(* IEC 61131-3 sources: bevling_machine/framework/sources/03_Units, 8 files *)

(* ---- FB_ClearanceUnit.st ---- *)
(* 模块说明：并行执行 P/Q 两路避让；两路都完成才继续，任一路故障向主流程报告。 *)
FUNCTION_BLOCK FB_ClearanceUnit
VAR_INPUT
    xExecute : BOOL; (* 子流程执行许可；须保持到完成，清 FALSE 复位该流程步骤和错误。 *)
    stRecipe : ST_Recipe; (* 待校验配方或上层传入的运行配方，字段含义见 ST_Recipe。 *)
END_VAR
VAR_IN_OUT
    aCommand : ARRAY[1..17] OF ST_DeviceCommand; (* 统一设备请求数组 1..17；子流程写请求，设备管理器执行。 *)
    aStatus : ARRAY[1..17] OF ST_DeviceStatus; (* 各设备的反馈数组 1..17，供判断忙、完成序号、故障和位置。 *)
    udiCounter : UDINT; (* 全机共享的动作序号计数器，通过引用传递；由 F_NextID 分配，0 不使用。 *)
END_VAR
VAR_OUTPUT
    xDone : BOOL; (* 本子流程完成标志；执行许可撤销后复位。 *)
    xError : BOOL; (* 本设备或本子流程发生故障；具体原因见对应错误码。 *)
    udiErrorID : UDINT; (* 错误码；0 表示无错误，设备或流程发生异常时赋值。 *)
    uiLengthStep : UINT; (* 定长支线当前步骤，供监控定位等待点。 *)
    uiTransferStep : UINT; (* 流利条/侧推/侧挡支线当前步骤，供监控定位等待点。 *)
END_VAR
VAR
    fbLength : FB_ClearLength; (* P 支线：D5 升起、D4 移开。 *)
    fbTransfer : FB_ClearTransfer; (* 切割前流利条/侧推/侧挡避让支线。 *)
END_VAR
FUNCTION_BLOCK FB_ClearanceUnit
(* P/Q 两路同一扫描使能；xDone 使用 AND，任一路未完成均不得继续。 *)
fbLength(xExecute:=xExecute,stRecipe:=stRecipe,aCommand:=aCommand,aStatus:=aStatus,udiCounter:=udiCounter);
fbTransfer(xExecute:=xExecute,stRecipe:=stRecipe,aCommand:=aCommand,aStatus:=aStatus,udiCounter:=udiCounter);
xDone := fbLength.xDone AND fbTransfer.xDone;
xError := fbLength.xError OR fbTransfer.xError;
udiErrorID := MAX(fbLength.udiErrorID,fbTransfer.udiErrorID);
uiLengthStep := fbLength.uiStep; uiTransferStep := fbTransfer.uiStep;

(* ---- FB_ClearLength.st ---- *)
(* 模块说明：切割前避让支线 P：D5 定长升起，再将 D4 移到避让位置。每步等待本次序号完成。 *)
FUNCTION_BLOCK FB_ClearLength
VAR_INPUT
    xExecute : BOOL; (* 子流程执行许可；须保持到完成，清 FALSE 复位该流程步骤和错误。 *)
    stRecipe : ST_Recipe; (* 待校验配方或上层传入的运行配方，字段含义见 ST_Recipe。 *)
END_VAR
VAR_IN_OUT
    aCommand : ARRAY[1..17] OF ST_DeviceCommand; (* 统一设备请求数组 1..17；子流程写请求，设备管理器执行。 *)
    aStatus : ARRAY[1..17] OF ST_DeviceStatus; (* 各设备的反馈数组 1..17，供判断忙、完成序号、故障和位置。 *)
    udiCounter : UDINT; (* 全机共享的动作序号计数器，通过引用传递；由 F_NextID 分配，0 不使用。 *)
END_VAR
VAR_OUTPUT
    xDone : BOOL; (* 本子流程完成标志；执行许可撤销后复位。 *)
    xError : BOOL; (* 本设备或本子流程发生故障；具体原因见对应错误码。 *)
    udiErrorID : UDINT; (* 非法步骤码 4100；动作超时码=4100+uiStep，可据此定位本支线等待点。 *)
    uiStep : UINT; (* 当前子步骤：0 待机，10/20/... 执行动作，1000 完成；切勿在线强制跳步。 *)
END_VAR
VAR
    uiPrevStep : UINT := 65535; (* 上扫描步骤，用于判断本扫描是否刚进入新步骤。 *)
    udiToken : UDINT; (* 本步骤专用动作序号；同一步中的设备共用该号，以排除旧完成信号。 *)
    xEntry : BOOL; (* 本扫描为新步骤入口；用于分配新序号并复位步骤超时计时。 *)
    tonStep : TON; (* 步骤超时定时器；进入新步骤时复位，超时错误码由模块及当前步号组成。 *)
    tonSpray : TON; (* 通用子流程模板的喷油定时器，只有 FB_ReturnKnife 用其完成条件。 *)
END_VAR
FUNCTION_BLOCK FB_ClearLength
(* 执行许可撤销即复位；步骤入口换新序号，每步等待本次动作完成，超时码=模块基码+步号。 *)
IF NOT xExecute THEN uiStep := 0; xError := FALSE; udiErrorID := 0; END_IF;
xEntry := uiStep <> uiPrevStep;
IF xEntry THEN udiToken := F_NextID(udiCounter); END_IF;
uiPrevStep := uiStep;
tonStep(IN := xExecute AND (uiStep > 0) AND (uiStep < 1000) AND NOT xEntry, PT := stRecipe.tStepTimeout);
tonSpray(IN := xExecute AND (uiStep = 10) AND aStatus[13].xActive, PT := stRecipe.tSpray);
IF xExecute AND NOT xError THEN
CASE uiStep OF
0: (* 待机；许可有效时进入首个动作。 *) uiStep := 10;
10: (* P010 定长 D5 升起避让；确认本次动作完成后再允许 D4 平移。 *)
aCommand[5] := F_Command(E_DeviceAction.Position, udiToken, 0.0, stRecipe.lrPositionVelocity);
IF F_Done(aStatus[5], udiToken) THEN uiStep := 20; END_IF;
20: (* P020 定长 D4 移到配方避让位置，等待本次序号完成。 *)
aCommand[4] := F_Command(E_DeviceAction.Position, udiToken, stRecipe.lrLengthClear, stRecipe.lrPositionVelocity);
IF F_Done(aStatus[4], udiToken) THEN uiStep := 1000; END_IF;
1000: (* 本支线完成，保持至 xExecute 撤销。 *) ;
ELSE xError := TRUE; udiErrorID := 4100;
END_CASE;
IF tonStep.Q THEN xError := TRUE; udiErrorID := 4100 + UINT_TO_UDINT(uiStep); END_IF;
END_IF;
xDone := xExecute AND (uiStep = 1000) AND NOT xError;

(* ---- FB_ClearTransfer.st ---- *)
(* 模块说明：切割前避让支线 Q：G4 流利条下降、G3 解除侧推、G2 侧挡下降。 *)
FUNCTION_BLOCK FB_ClearTransfer
VAR_INPUT
    xExecute : BOOL; (* 子流程执行许可；须保持到完成，清 FALSE 复位该流程步骤和错误。 *)
    stRecipe : ST_Recipe; (* 待校验配方或上层传入的运行配方，字段含义见 ST_Recipe。 *)
END_VAR
VAR_IN_OUT
    aCommand : ARRAY[1..17] OF ST_DeviceCommand; (* 统一设备请求数组 1..17；子流程写请求，设备管理器执行。 *)
    aStatus : ARRAY[1..17] OF ST_DeviceStatus; (* 各设备的反馈数组 1..17，供判断忙、完成序号、故障和位置。 *)
    udiCounter : UDINT; (* 全机共享的动作序号计数器，通过引用传递；由 F_NextID 分配，0 不使用。 *)
END_VAR
VAR_OUTPUT
    xDone : BOOL; (* 本子流程完成标志；执行许可撤销后复位。 *)
    xError : BOOL; (* 本设备或本子流程发生故障；具体原因见对应错误码。 *)
    udiErrorID : UDINT; (* 非法步骤码 4200；动作超时码=4200+uiStep，可据此定位本支线等待点。 *)
    uiStep : UINT; (* 当前子步骤：0 待机，10/20/... 执行动作，1000 完成；切勿在线强制跳步。 *)
END_VAR
VAR
    uiPrevStep : UINT := 65535; (* 上扫描步骤，用于判断本扫描是否刚进入新步骤。 *)
    udiToken : UDINT; (* 本步骤专用动作序号；同一步中的设备共用该号，以排除旧完成信号。 *)
    xEntry : BOOL; (* 本扫描为新步骤入口；用于分配新序号并复位步骤超时计时。 *)
    tonStep : TON; (* 步骤超时定时器；进入新步骤时复位，超时错误码由模块及当前步号组成。 *)
    tonSpray : TON; (* 通用子流程模板的喷油定时器，只有 FB_ReturnKnife 用其完成条件。 *)
END_VAR
FUNCTION_BLOCK FB_ClearTransfer
(* 执行许可撤销即复位；步骤入口换新序号，每步等待本次动作完成，超时码=模块基码+步号。 *)
IF NOT xExecute THEN uiStep := 0; xError := FALSE; udiErrorID := 0; END_IF;
xEntry := uiStep <> uiPrevStep;
IF xEntry THEN udiToken := F_NextID(udiCounter); END_IF;
uiPrevStep := uiStep;
tonStep(IN := xExecute AND (uiStep > 0) AND (uiStep < 1000) AND NOT xEntry, PT := stRecipe.tStepTimeout);
tonSpray(IN := xExecute AND (uiStep = 10) AND aStatus[13].xActive, PT := stRecipe.tSpray);
IF xExecute AND NOT xError THEN
CASE uiStep OF
0: (* 待机；许可有效时进入首个动作。 *) uiStep := 10;
10: (* Q010 流利条 G4 下降。 *)
aCommand[12] := F_Command(E_DeviceAction.Position, udiToken, 0.0, stRecipe.lrPositionVelocity);
IF F_Done(aStatus[12], udiToken) THEN uiStep := 20; END_IF;
20: (* Q020 推动气缸 G3 放开。 *)
aCommand[11] := F_Command(E_DeviceAction.Position, udiToken, 0.0, stRecipe.lrPositionVelocity);
IF F_Done(aStatus[11], udiToken) THEN uiStep := 30; END_IF;
30: (* Q030 侧挡 G2 下降。目标固定发 1.0：本层不知道侧挡是单缸还是 300/450/600 三缸组，
   由设备层自己解释——仿真气缸按 1.0 到伸出端，真实三缸组按当前料型选缸下降。 *)
aCommand[10] := F_Command(E_DeviceAction.Position, udiToken, 1.0, stRecipe.lrPositionVelocity);
IF F_Done(aStatus[10], udiToken) THEN uiStep := 1000; END_IF;
1000: (* 本支线完成，保持至 xExecute 撤销。 *) ;
ELSE xError := TRUE; udiErrorID := 4200;
END_CASE;
IF tonStep.Q THEN xError := TRUE; udiErrorID := 4200 + UINT_TO_UDINT(uiStep); END_IF;
END_IF;
xDone := xExecute AND (uiStep = 1000) AND NOT xError;

(* ---- FB_Initialize.st ---- *)
(* 模块说明：初始姿态整理流程。20 步摆好避让姿态后，25 步让真实轴回零，30 步再按配方绝对定位。 *)
FUNCTION_BLOCK FB_Initialize
VAR_INPUT
    xExecute : BOOL; (* 子流程执行许可；须保持到完成，清 FALSE 复位该流程步骤和错误。 *)
    stRecipe : ST_Recipe; (* 待校验配方或上层传入的运行配方，字段含义见 ST_Recipe。 *)
END_VAR
VAR_IN_OUT
    aCommand : ARRAY[1..17] OF ST_DeviceCommand; (* 统一设备请求数组 1..17；子流程写请求，设备管理器执行。 *)
    aStatus : ARRAY[1..17] OF ST_DeviceStatus; (* 各设备的反馈数组 1..17，供判断忙、完成序号、故障和位置。 *)
    udiCounter : UDINT; (* 全机共享的动作序号计数器，通过引用传递；由 F_NextID 分配，0 不使用。 *)
END_VAR
VAR_OUTPUT
    xDone : BOOL; (* 本子流程完成标志；执行许可撤销后复位。 *)
    xError : BOOL; (* 本设备或本子流程发生故障；具体原因见对应错误码。 *)
    udiErrorID : UDINT; (* 非法步骤码 4600；动作超时码=4600+uiStep，可据此定位本支线等待点。 *)
    uiStep : UINT; (* 当前子步骤：0 待机，10/20/25/30/40 执行动作，1000 完成；切勿在线强制跳步。 *)
END_VAR
VAR
    uiPrevStep : UINT := 65535; (* 上扫描步骤，用于判断本扫描是否刚进入新步骤。 *)
    udiToken : UDINT; (* 本步骤专用动作序号；同一步中的设备共用该号，以排除旧完成信号。 *)
    xEntry : BOOL; (* 本扫描为新步骤入口；用于分配新序号并复位步骤超时计时。 *)
    tonStep : TON; (* 步骤超时定时器；进入新步骤时复位，超时错误码由模块及当前步号组成。 *)
    tonSpray : TON; (* 通用子流程模板的喷油定时器，只有 FB_ReturnKnife 用其完成条件。 *)
END_VAR
FUNCTION_BLOCK FB_Initialize
(* 执行许可撤销即复位；步骤入口换新序号，每步等待本次动作完成，超时码=模块基码+步号。 *)
IF NOT xExecute THEN uiStep := 0; xError := FALSE; udiErrorID := 0; END_IF;
xEntry := uiStep <> uiPrevStep;
IF xEntry THEN udiToken := F_NextID(udiCounter); END_IF;
uiPrevStep := uiStep;
tonStep(IN := xExecute AND (uiStep > 0) AND (uiStep < 1000) AND NOT xEntry, PT := stRecipe.tStepTimeout);
tonSpray(IN := xExecute AND (uiStep = 10) AND aStatus[13].xActive, PT := stRecipe.tSpray);
IF xExecute AND NOT xError THEN
CASE uiStep OF
0: (* 待机；许可有效时进入首个动作。 *) uiStep := 10;
10: (* 仿真初始化 10：同时抬起 G9、抬起 G1、打开 G8，三项都完成才继续。 *)
aCommand[17] := F_Command(E_DeviceAction.Position, udiToken, 0.0, stRecipe.lrPositionVelocity);
aCommand[9] := F_Command(E_DeviceAction.Position, udiToken, 0.0, stRecipe.lrPositionVelocity);
aCommand[16] := F_Command(E_DeviceAction.Position, udiToken, 0.0, stRecipe.lrPositionVelocity);
IF F_Done(aStatus[17], udiToken) AND F_Done(aStatus[9], udiToken) AND F_Done(aStatus[16], udiToken) THEN uiStep := 20; END_IF;
20: (* 仿真初始化 20：D5 升起、G2 提升、G3 释放、G4 提升、G7 下降，全部完成再定位。 *)
aCommand[5] := F_Command(E_DeviceAction.Position, udiToken, 0.0, stRecipe.lrPositionVelocity);
aCommand[10] := F_Command(E_DeviceAction.Position, udiToken, 0.0, stRecipe.lrPositionVelocity);
aCommand[11] := F_Command(E_DeviceAction.Position, udiToken, 0.0, stRecipe.lrPositionVelocity);
aCommand[12] := F_Command(E_DeviceAction.Position, udiToken, 1.0, stRecipe.lrPositionVelocity);
aCommand[15] := F_Command(E_DeviceAction.Position, udiToken, 0.0, stRecipe.lrPositionVelocity);
IF F_Done(aStatus[5], udiToken) AND F_Done(aStatus[10], udiToken) AND F_Done(aStatus[11], udiToken) AND F_Done(aStatus[12], udiToken) AND F_Done(aStatus[15], udiToken) THEN uiStep := 25; END_IF;
25: (* 初始化 25：真实轴回零。D2 走刀与 D8 旋转是真轴，D4 定长平移当前为仿真，由仿真在 tSimAction 后完成。
       D3 盘刀是连续旋转主轴，自动流程只下发 Run 不定位，因此不参与回零，也不占本步完成条件。 *)
aCommand[2] := F_Command(E_DeviceAction.Home, udiToken, 0.0, 0.0);
aCommand[4] := F_Command(E_DeviceAction.Home, udiToken, 0.0, 0.0);
aCommand[8] := F_Command(E_DeviceAction.Home, udiToken, 0.0, 0.0);
IF F_Done(aStatus[2], udiToken) AND F_Done(aStatus[4], udiToken) AND F_Done(aStatus[8], udiToken) THEN uiStep := 30; END_IF;
30: (* 仿真初始化 30：D2/D4/D7/D8 移至示例初始坐标，全部完成才继续。 *)
aCommand[2] := F_Command(E_DeviceAction.Position, udiToken, stRecipe.lrCutHome, stRecipe.lrPositionVelocity);
aCommand[4] := F_Command(E_DeviceAction.Position, udiToken, stRecipe.lrLengthPosition, stRecipe.lrPositionVelocity);
aCommand[7] := F_Command(E_DeviceAction.Position, udiToken, stRecipe.lrGripperHome, stRecipe.lrPositionVelocity);
aCommand[8] := F_Command(E_DeviceAction.Position, udiToken, 0.0, stRecipe.lrPositionVelocity);
IF F_Done(aStatus[2], udiToken) AND F_Done(aStatus[4], udiToken) AND F_Done(aStatus[7], udiToken) AND F_Done(aStatus[8], udiToken) THEN uiStep := 40; END_IF;
40: (* 仿真初始化 40：D5 下降，准备进入来料检测。 *)
aCommand[5] := F_Command(E_DeviceAction.Position, udiToken, 1.0, stRecipe.lrPositionVelocity);
IF F_Done(aStatus[5], udiToken) THEN uiStep := 1000; END_IF;
1000: (* 本支线完成，保持至 xExecute 撤销。 *) ;
ELSE xError := TRUE; udiErrorID := 4600;
END_CASE;
IF tonStep.Q THEN xError := TRUE; udiErrorID := 4600 + UINT_TO_UDINT(uiStep); END_IF;
END_IF;
xDone := xExecute AND (uiStep = 1000) AND NOT xError;

(* ---- FB_PostCut.st ---- *)
(* 模块说明：切割后先 G9 抬刀，再 G1 抬压；之后同时执行回刀、机械手移料、定长复位，三路全完成才结束。 *)
FUNCTION_BLOCK FB_PostCut
VAR_INPUT
    xExecute : BOOL; (* 子流程执行许可；须保持到完成，清 FALSE 复位该流程步骤和错误。 *)
    stRecipe : ST_Recipe; (* 待校验配方或上层传入的运行配方，字段含义见 ST_Recipe。 *)
END_VAR
VAR_IN_OUT
    aCommand : ARRAY[1..17] OF ST_DeviceCommand; (* 统一设备请求数组 1..17；子流程写请求，设备管理器执行。 *)
    aStatus : ARRAY[1..17] OF ST_DeviceStatus; (* 各设备的反馈数组 1..17，供判断忙、完成序号、故障和位置。 *)
    udiCounter : UDINT; (* 全机共享的动作序号计数器，通过引用传递；由 F_NextID 分配，0 不使用。 *)
END_VAR
VAR_OUTPUT
    xDone : BOOL; (* 本子流程完成标志；执行许可撤销后复位。 *)
    xError : BOOL; (* 本设备或本子流程发生故障；具体原因见对应错误码。 *)
    udiErrorID : UDINT; (* 非法总步骤为 4700，超时为 4700+总步号；支线故障则向上传递支线错误码。 *)
    uiStep : UINT; (* 当前子步骤：0 待机，10/20/... 执行动作，1000 完成；切勿在线强制跳步。 *)
    uiKnifeStep : UINT; (* 收尾回刀支线 A 当前步骤：喷油、回刀或完成。 *)
    uiUnloadStep : UINT; (* 机械手移料支线 B 步骤，10..110 每步加 10，1000 完成；详见 FB_Unload。 *)
    uiLengthStep : UINT; (* 定长支线当前步骤，供监控定位等待点。 *)
END_VAR
VAR
    fbKnife : FB_ReturnKnife; (* 收尾支线 A：喷油后回刀。 *)
    fbUnload : FB_Unload; (* 收尾支线 B：机械手移料，含后退、下降、最终回位。 *)
    fbLength : FB_ResetLength; (* C 支线：D4 回检测位置、D5 下降、确认下降到位。 *)
    uiPrevStep : UINT := 65535; (* 上扫描步骤，用于判断本扫描是否刚进入新步骤。 *)
    udiToken : UDINT; (* 本步骤专用动作序号；同一步中的设备共用该号，以排除旧完成信号。 *)
    xEntry : BOOL; (* 本扫描为新步骤入口；用于分配新序号并复位步骤超时计时。 *)
    tonStep : TON; (* 步骤超时定时器；进入新步骤时复位，超时错误码由模块及当前步号组成。 *)
END_VAR
FUNCTION_BLOCK FB_PostCut
IF NOT xExecute THEN uiStep := 0; xError := FALSE; udiErrorID := 0; END_IF
(* 每个总步骤分配新序号；等待三路期间保留总步骤超时。 *)
xEntry := uiStep <> uiPrevStep;
IF xEntry THEN udiToken := F_NextID(udiCounter); END_IF
uiPrevStep := uiStep;
tonStep(IN:=xExecute AND NOT xEntry AND (uiStep>0) AND (uiStep<1000),PT:=stRecipe.tStepTimeout);
IF xExecute AND NOT xError THEN
    CASE uiStep OF
    0: (* 待机，执行许可有效后进入抬刀。 *) uiStep := 10;
    10: (* 先 G9 盘刀提升；同时保持 G1 下压，刀没抬起来之前不能松压板。 *)
        aCommand[9] := F_Command(E_DeviceAction.Position,udiToken,1.0,stRecipe.lrPositionVelocity);
        aCommand[17] := F_Command(E_DeviceAction.Position,udiToken,0.0,stRecipe.lrPositionVelocity);
        IF F_Done(aStatus[17],udiToken) THEN uiStep := 20; END_IF
    20: (* 再 G1 下压提升，等待本次序号完成。 *)
        aCommand[9] := F_Command(E_DeviceAction.Position,udiToken,0.0,stRecipe.lrPositionVelocity);
        IF F_Done(aStatus[9],udiToken) THEN uiStep := 30; END_IF
    30: (* 等待回刀、机械手移料、定长复位三路全部完成。 *)
        IF fbKnife.xDone AND fbUnload.xDone AND fbLength.xDone THEN uiStep := 1000; END_IF
    1000: (* 三路收尾结束，保持完成反馈直到执行许可撤销。 *) ;
    ELSE xError := TRUE; udiErrorID := 4700;
    END_CASE
    IF tonStep.Q THEN xError := TRUE; udiErrorID := 4700+UINT_TO_UDINT(uiStep); END_IF
END_IF
(* 三路只在总步骤 30 同时使能，并且每扫描调用；等待三路全完成才退出。 *)
fbKnife(xExecute:=xExecute AND (uiStep=30),stRecipe:=stRecipe,aCommand:=aCommand,aStatus:=aStatus,udiCounter:=udiCounter);
fbUnload(xExecute:=xExecute AND (uiStep=30),stRecipe:=stRecipe,aCommand:=aCommand,aStatus:=aStatus,udiCounter:=udiCounter);
fbLength(xExecute:=xExecute AND (uiStep=30),stRecipe:=stRecipe,aCommand:=aCommand,aStatus:=aStatus,udiCounter:=udiCounter);
IF fbKnife.xError OR fbUnload.xError OR fbLength.xError THEN
    xError:=TRUE; udiErrorID:=MAX(fbKnife.udiErrorID,MAX(fbUnload.udiErrorID,fbLength.udiErrorID));
END_IF
xDone := xExecute AND (uiStep=1000) AND NOT xError;
uiKnifeStep:=fbKnife.uiStep; uiUnloadStep:=fbUnload.uiStep; uiLengthStep:=fbLength.uiStep;

(* ---- FB_ResetLength.st ---- *)
(* 模块说明：收尾支线 C：D4 回检测位置、D5 下降到位、确认下降位置；随后具备来料检测条件。 *)
FUNCTION_BLOCK FB_ResetLength
VAR_INPUT
    xExecute : BOOL; (* 子流程执行许可；须保持到完成，清 FALSE 复位该流程步骤和错误。 *)
    stRecipe : ST_Recipe; (* 待校验配方或上层传入的运行配方，字段含义见 ST_Recipe。 *)
END_VAR
VAR_IN_OUT
    aCommand : ARRAY[1..17] OF ST_DeviceCommand; (* 统一设备请求数组 1..17；子流程写请求，设备管理器执行。 *)
    aStatus : ARRAY[1..17] OF ST_DeviceStatus; (* 各设备的反馈数组 1..17，供判断忙、完成序号、故障和位置。 *)
    udiCounter : UDINT; (* 全机共享的动作序号计数器，通过引用传递；由 F_NextID 分配，0 不使用。 *)
END_VAR
VAR_OUTPUT
    xDone : BOOL; (* 本子流程完成标志；执行许可撤销后复位。 *)
    xError : BOOL; (* 本设备或本子流程发生故障；具体原因见对应错误码。 *)
    udiErrorID : UDINT; (* 非法步骤码 4500；动作超时码=4500+uiStep，可据此定位本支线等待点。 *)
    uiStep : UINT; (* 当前子步骤：0 待机，10/20/... 执行动作，1000 完成；切勿在线强制跳步。 *)
END_VAR
VAR
    uiPrevStep : UINT := 65535; (* 上扫描步骤，用于判断本扫描是否刚进入新步骤。 *)
    udiToken : UDINT; (* 本步骤专用动作序号；同一步中的设备共用该号，以排除旧完成信号。 *)
    xEntry : BOOL; (* 本扫描为新步骤入口；用于分配新序号并复位步骤超时计时。 *)
    tonStep : TON; (* 步骤超时定时器；进入新步骤时复位，超时错误码由模块及当前步号组成。 *)
    tonSpray : TON; (* 通用子流程模板的喷油定时器，只有 FB_ReturnKnife 用其完成条件。 *)
END_VAR
FUNCTION_BLOCK FB_ResetLength
(* 执行许可撤销即复位；步骤入口换新序号，每步等待本次动作完成，超时码=模块基码+步号。 *)
IF NOT xExecute THEN uiStep := 0; xError := FALSE; udiErrorID := 0; END_IF;
xEntry := uiStep <> uiPrevStep;
IF xEntry THEN udiToken := F_NextID(udiCounter); END_IF;
uiPrevStep := uiStep;
tonStep(IN := xExecute AND (uiStep > 0) AND (uiStep < 1000) AND NOT xEntry, PT := stRecipe.tStepTimeout);
tonSpray(IN := xExecute AND (uiStep = 10) AND aStatus[13].xActive, PT := stRecipe.tSpray);
IF xExecute AND NOT xError THEN
CASE uiStep OF
0: (* 待机；许可有效时进入首个动作。 *) uiStep := 10;
10: (* C010 定长 D4 回到配方检测位置 lrLengthPosition。 *)
aCommand[4] := F_Command(E_DeviceAction.Position, udiToken, stRecipe.lrLengthPosition, stRecipe.lrPositionVelocity);
IF F_Done(aStatus[4], udiToken) THEN uiStep := 20; END_IF;
20: (* C020 D4 到位后，定长 D5 下降。 *)
aCommand[5] := F_Command(E_DeviceAction.Position, udiToken, 1.0, stRecipe.lrPositionVelocity);
IF F_Done(aStatus[5], udiToken) THEN uiStep := 30; END_IF;
30: (* C030 确认 D5 下降端到位，后续送料才具备光电检测条件。 *)
IF F_At(aStatus[5],1.0) THEN uiStep := 1000; END_IF;
1000: (* 本支线完成，保持至 xExecute 撤销。 *) ;
ELSE xError := TRUE; udiErrorID := 4500;
END_CASE;
IF tonStep.Q THEN xError := TRUE; udiErrorID := 4500 + UINT_TO_UDINT(uiStep); END_IF;
END_IF;
xDone := xExecute AND (uiStep = 1000) AND NOT xError;

(* ---- FB_ReturnKnife.st ---- *)
(* 模块说明：收尾支线 A：G5 喷油到设定时间，再令 D2 回刀。喷油仅在第一步保持请求。 *)
FUNCTION_BLOCK FB_ReturnKnife
VAR_INPUT
    xExecute : BOOL; (* 子流程执行许可；须保持到完成，清 FALSE 复位该流程步骤和错误。 *)
    stRecipe : ST_Recipe; (* 待校验配方或上层传入的运行配方，字段含义见 ST_Recipe。 *)
END_VAR
VAR_IN_OUT
    aCommand : ARRAY[1..17] OF ST_DeviceCommand; (* 统一设备请求数组 1..17；子流程写请求，设备管理器执行。 *)
    aStatus : ARRAY[1..17] OF ST_DeviceStatus; (* 各设备的反馈数组 1..17，供判断忙、完成序号、故障和位置。 *)
    udiCounter : UDINT; (* 全机共享的动作序号计数器，通过引用传递；由 F_NextID 分配，0 不使用。 *)
END_VAR
VAR_OUTPUT
    xDone : BOOL; (* 本子流程完成标志；执行许可撤销后复位。 *)
    xError : BOOL; (* 本设备或本子流程发生故障；具体原因见对应错误码。 *)
    udiErrorID : UDINT; (* 非法步骤码 4300；动作超时码=4300+uiStep，可据此定位本支线等待点。 *)
    uiStep : UINT; (* 当前子步骤：0 待机，10/20/... 执行动作，1000 完成；切勿在线强制跳步。 *)
END_VAR
VAR
    uiPrevStep : UINT := 65535; (* 上扫描步骤，用于判断本扫描是否刚进入新步骤。 *)
    udiToken : UDINT; (* 本步骤专用动作序号；同一步中的设备共用该号，以排除旧完成信号。 *)
    xEntry : BOOL; (* 本扫描为新步骤入口；用于分配新序号并复位步骤超时计时。 *)
    tonStep : TON; (* 步骤超时定时器；进入新步骤时复位，超时错误码由模块及当前步号组成。 *)
    tonSpray : TON; (* 通用子流程模板的喷油定时器，只有 FB_ReturnKnife 用其完成条件。 *)
END_VAR
FUNCTION_BLOCK FB_ReturnKnife
(* 执行许可撤销即复位；步骤入口换新序号，每步等待本次动作完成，超时码=模块基码+步号。 *)
IF NOT xExecute THEN uiStep := 0; xError := FALSE; udiErrorID := 0; END_IF;
xEntry := uiStep <> uiPrevStep;
IF xEntry THEN udiToken := F_NextID(udiCounter); END_IF;
uiPrevStep := uiStep;
tonStep(IN := xExecute AND (uiStep > 0) AND (uiStep < 1000) AND NOT xEntry, PT := stRecipe.tStepTimeout);
tonSpray(IN := xExecute AND (uiStep = 10) AND aStatus[13].xActive, PT := stRecipe.tSpray);
IF xExecute AND NOT xError THEN
CASE uiStep OF
0: (* 待机；许可有效时进入首个动作。 *) uiStep := 10;
10: (* A010 G5 喷油并等待 tSpray；喷油建立后才开始计时。 *)
aCommand[13] := F_Command(E_DeviceAction.Run, udiToken, 0.0, 0.0);
IF tonSpray.Q THEN uiStep := 20; END_IF;
20: (* A020 结束喷油请求，D2 回到 lrCutHome，等待到位。 *)
aCommand[2] := F_Command(E_DeviceAction.Position, udiToken, stRecipe.lrCutHome, stRecipe.lrReturnVelocity);
IF F_Done(aStatus[2], udiToken) THEN uiStep := 1000; END_IF;
1000: (* 本支线完成，保持至 xExecute 撤销。 *) ;
ELSE xError := TRUE; udiErrorID := 4300;
END_CASE;
IF tonStep.Q THEN xError := TRUE; udiErrorID := 4300 + UINT_TO_UDINT(uiStep); END_IF;
END_IF;
xDone := xExecute AND (uiStep = 1000) AND NOT xError;

(* ---- FB_Unload.st ---- *)
(* 模块说明：收尾支线 B：机械手移料。后退、下降、最终回位是三个独立动作，全部完成后才允许下一轮送料。 *)
FUNCTION_BLOCK FB_Unload
VAR_INPUT
    xExecute : BOOL; (* 子流程执行许可；须保持到完成，清 FALSE 复位该流程步骤和错误。 *)
    stRecipe : ST_Recipe; (* 待校验配方或上层传入的运行配方，字段含义见 ST_Recipe。 *)
END_VAR
VAR_IN_OUT
    aCommand : ARRAY[1..17] OF ST_DeviceCommand; (* 统一设备请求数组 1..17；子流程写请求，设备管理器执行。 *)
    aStatus : ARRAY[1..17] OF ST_DeviceStatus; (* 各设备的反馈数组 1..17，供判断忙、完成序号、故障和位置。 *)
    udiCounter : UDINT; (* 全机共享的动作序号计数器，通过引用传递；由 F_NextID 分配，0 不使用。 *)
END_VAR
VAR_OUTPUT
    xDone : BOOL; (* 本子流程完成标志；执行许可撤销后复位。 *)
    xError : BOOL; (* 本设备或本子流程发生故障；具体原因见对应错误码。 *)
    udiErrorID : UDINT; (* 非法步骤码 4400；动作超时码=4400+uiStep，可据此定位本支线等待点。 *)
    uiStep : UINT; (* 当前子步骤：0 待机，10/20/... 执行动作，1000 完成；切勿在线强制跳步。 *)
END_VAR
VAR
    uiPrevStep : UINT := 65535; (* 上扫描步骤，用于判断本扫描是否刚进入新步骤。 *)
    udiToken : UDINT; (* 本步骤专用动作序号；同一步中的设备共用该号，以排除旧完成信号。 *)
    xEntry : BOOL; (* 本扫描为新步骤入口；用于分配新序号并复位步骤超时计时。 *)
    tonStep : TON; (* 步骤超时定时器；进入新步骤时复位，超时错误码由模块及当前步号组成。 *)
    tonSpray : TON; (* 通用子流程模板的喷油定时器，只有 FB_ReturnKnife 用其完成条件。 *)
END_VAR
FUNCTION_BLOCK FB_Unload
(* 执行许可撤销即复位；步骤入口换新序号，每步等待本次动作完成，超时码=模块基码+步号。 *)
IF NOT xExecute THEN uiStep := 0; xError := FALSE; udiErrorID := 0; END_IF;
xEntry := uiStep <> uiPrevStep;
IF xEntry THEN udiToken := F_NextID(udiCounter); END_IF;
uiPrevStep := uiStep;
tonStep(IN := xExecute AND (uiStep > 0) AND (uiStep < 1000) AND NOT xEntry, PT := stRecipe.tStepTimeout);
tonSpray(IN := xExecute AND (uiStep = 10) AND aStatus[13].xActive, PT := stRecipe.tSpray);
IF xExecute AND NOT xError THEN
CASE uiStep OF
0: (* 待机；许可有效时进入首个动作。 *) uiStep := 10;
10: (* B010 侧挡 G2 提升。 *)
aCommand[10] := F_Command(E_DeviceAction.Position, udiToken, 0.0, stRecipe.lrPositionVelocity);
IF F_Done(aStatus[10], udiToken) THEN uiStep := 20; END_IF;
20: (* B020 流利条 G4 提升。 *)
aCommand[12] := F_Command(E_DeviceAction.Position, udiToken, 1.0, stRecipe.lrPositionVelocity);
IF F_Done(aStatus[12], udiToken) THEN uiStep := 30; END_IF;
30: (* B030 机械手 G7 提升。 *)
aCommand[15] := F_Command(E_DeviceAction.Position, udiToken, 1.0, stRecipe.lrPositionVelocity);
IF F_Done(aStatus[15], udiToken) THEN uiStep := 40; END_IF;
40: (* B040 夹爪 G8 打开，准备前进取料。 *)
aCommand[16] := F_Command(E_DeviceAction.Position, udiToken, 0.0, stRecipe.lrPositionVelocity);
IF F_Done(aStatus[16], udiToken) THEN uiStep := 50; END_IF;
50: (* B050 机械手 D7 前进到取料位置 lrGripperFront。 *)
aCommand[7] := F_Command(E_DeviceAction.Position, udiToken, stRecipe.lrGripperFront, stRecipe.lrPositionVelocity);
IF F_Done(aStatus[7], udiToken) THEN uiStep := 60; END_IF;
60: (* B060 夹爪 G8 夹紧，确认后才拉料。 *)
aCommand[16] := F_Command(E_DeviceAction.Position, udiToken, 1.0, stRecipe.lrPositionVelocity);
IF F_Done(aStatus[16], udiToken) THEN uiStep := 70; END_IF;
70: (* B070 机械手 D7 拉料到 lrGripperPull。 *)
aCommand[7] := F_Command(E_DeviceAction.Position, udiToken, stRecipe.lrGripperPull, stRecipe.lrPositionVelocity);
IF F_Done(aStatus[7], udiToken) THEN uiStep := 80; END_IF;
80: (* B080 夹爪 G8 打开，释放移走的料。 *)
aCommand[16] := F_Command(E_DeviceAction.Position, udiToken, 0.0, stRecipe.lrPositionVelocity);
IF F_Done(aStatus[16], udiToken) THEN uiStep := 90; END_IF;
90: (* B090 保持机械手抬升，D7 后退至 lrGripperBack；此时不是最终回位。 *)
aCommand[7] := F_Command(E_DeviceAction.Position, udiToken, stRecipe.lrGripperBack, stRecipe.lrPositionVelocity);
IF F_Done(aStatus[7], udiToken) THEN uiStep := 100; END_IF;
100: (* B100 后退到位后，G7 下降。 *)
aCommand[15] := F_Command(E_DeviceAction.Position, udiToken, 0.0, stRecipe.lrPositionVelocity);
IF F_Done(aStatus[15], udiToken) THEN uiStep := 110; END_IF;
110: (* B110 下降到位后，D7 再回 lrGripperHome；本支线结束前不允许送料。 *)
aCommand[7] := F_Command(E_DeviceAction.Position, udiToken, stRecipe.lrGripperHome, stRecipe.lrPositionVelocity);
IF F_Done(aStatus[7], udiToken) THEN uiStep := 1000; END_IF;
1000: (* 本支线完成，保持至 xExecute 撤销。 *) ;
ELSE xError := TRUE; udiErrorID := 4400;
END_CASE;
IF tonStep.Q THEN xError := TRUE; udiErrorID := 4400 + UINT_TO_UDINT(uiStep); END_IF;
END_IF;
xDone := xExecute AND (uiStep = 1000) AND NOT xError;
